(* IEC 61131-3 sources: plc-vscode/tests/st/test-ready/trust-platform/examples/OSCAT/water_booster_pump_station/oop/src, 3 files *)

(* ---- Main.st ---- *)
(* Pattern role: IPump is the contract boundary for the Mediator and Observer example. *)
INTERFACE IPump EXTENDS IComponent
    PROPERTY PumpId : INT
    GET
    END_GET
    END_PROPERTY

    PROPERTY IsHealthy : BOOL
    GET
    END_GET
    END_PROPERTY

    PROPERTY IsRunning : BOOL
    GET
    END_GET
    END_PROPERTY

    PROPERTY RuntimeHours : REAL
    GET
    END_GET
    END_PROPERTY

    PROPERTY SpeedReference : REAL
    GET
    END_GET
    END_PROPERTY

    METHOD Run
    VAR_INPUT
        SpeedReference : REAL;
    END_VAR
    END_METHOD

    METHOD Stop
    END_METHOD
END_INTERFACE

(* Pattern role: IAlarmSubscriber is the contract boundary for the Mediator and Observer example. *)
INTERFACE IAlarmSubscriber
    METHOD OnAlarm
    VAR_INPUT
        ClassId : BYTE;
        Code : DWORD;
        SourceId : INT;
    END_VAR
    END_METHOD
END_INTERFACE

(* Pattern role: PumpDrive is a concrete implementation in the Mediator and Observer example. *)
FUNCTION_BLOCK PumpDrive IMPLEMENTS IPump
VAR
    IdValue : INT;
    FaultValue : BOOL;
    RemoteValue : BOOL := TRUE;
    RunningValue : BOOL;
    RuntimeValue : REAL;
    SpeedValue : REAL;
    ReadyValue : BOOL;
    ErrorValue : BOOL;
    ErrorIdValue : WORD;
    StatusValue : BYTE;
    RuntimeMeter : OntimeMeter;
END_VAR

METHOD PUBLIC Configure
VAR_INPUT
    PumpId : INT;
    RuntimeHoursInitial : REAL;
    Faulted : BOOL;
END_VAR
IdValue := PumpId;
RuntimeValue := RuntimeHoursInitial;
FaultValue := Faulted;
END_METHOD

METHOD PUBLIC Initialize
ReadyValue := TRUE;
RuntimeMeter.Initialize();
RuntimeMeter.Reset();
ClearError();
END_METHOD

METHOD PUBLIC Reset
RunningValue := FALSE;
SpeedValue := REAL#0.0;
ClearError();
END_METHOD

METHOD PUBLIC ClearError
ErrorValue := FALSE;
ErrorIdValue := WORD#0;
StatusValue := BYTE#0;
END_METHOD

METHOD PUBLIC Snapshot : ComponentStatus
VAR
    Result : ComponentStatus;
END_VAR
Result.Ready := ReadyValue;
Result.Error := ErrorValue;
Result.ErrorId := ErrorIdValue;
Result.Status := StatusValue;
Snapshot := Result;
END_METHOD

METHOD PUBLIC Run
VAR_INPUT
    SpeedReference : REAL;
END_VAR
IF NOT FaultValue AND RemoteValue THEN
    RunningValue := TRUE;
    SpeedValue := LIMIT(REAL#0.0, SpeedReference, REAL#100.0);
ELSE
    RunningValue := FALSE;
    SpeedValue := REAL#0.0;
END_IF;
RuntimeMeter.Update(Input := RunningValue);
END_METHOD

METHOD PUBLIC Stop
RunningValue := FALSE;
SpeedValue := REAL#0.0;
RuntimeMeter.Update(Input := FALSE);
END_METHOD

PUBLIC PROPERTY PumpId : INT
GET
    PumpId := IdValue;
END_GET
END_PROPERTY

PUBLIC PROPERTY IsHealthy : BOOL
GET
    IsHealthy := NOT FaultValue AND RemoteValue;
END_GET
END_PROPERTY

PUBLIC PROPERTY IsRunning : BOOL
GET
    IsRunning := RunningValue;
END_GET
END_PROPERTY

PUBLIC PROPERTY RuntimeHours : REAL
GET
    RuntimeHours := RuntimeValue;
END_GET
END_PROPERTY

PUBLIC PROPERTY SpeedReference : REAL
GET
    SpeedReference := SpeedValue;
END_GET
END_PROPERTY

PUBLIC PROPERTY Ready : BOOL
GET
    Ready := ReadyValue;
END_GET
END_PROPERTY

PUBLIC PROPERTY Error : BOOL
GET
    Error := ErrorValue;
END_GET
END_PROPERTY

PUBLIC PROPERTY ErrorId : WORD
GET
    ErrorId := ErrorIdValue;
END_GET
END_PROPERTY

PUBLIC PROPERTY Status : BYTE
GET
    Status := StatusValue;
END_GET
END_PROPERTY
END_FUNCTION_BLOCK

(* Pattern role: HistorianAlarmSubscriber is a concrete implementation in the Mediator and Observer example. *)
FUNCTION_BLOCK HistorianAlarmSubscriber IMPLEMENTS IAlarmSubscriber
VAR
    LastCodeValue : DWORD;
    CountValue : INT;
    Journal : DwordFifo32;
END_VAR

METHOD PUBLIC Initialize
Journal.Initialize();
Journal.Reset();
LastCodeValue := DWORD#0;
CountValue := INT#0;
END_METHOD

METHOD PUBLIC OnAlarm
VAR_INPUT
    ClassId : BYTE;
    Code : DWORD;
    SourceId : INT;
END_VAR
LastCodeValue := Code;
CountValue := CountValue + INT#1;
IF Journal.Push(Value := Code) THEN
END_IF;
END_METHOD

PUBLIC PROPERTY Count : INT
GET
    Count := CountValue;
END_GET
END_PROPERTY

PUBLIC PROPERTY LastCode : DWORD
GET
    LastCode := LastCodeValue;
END_GET
END_PROPERTY
END_FUNCTION_BLOCK

(* Pattern role: MqttAlarmSubscriber is a concrete implementation in the Mediator and Observer example. *)
FUNCTION_BLOCK MqttAlarmSubscriber IMPLEMENTS IAlarmSubscriber
VAR
    PublishReadyValue : BOOL;
    LastCodeValue : DWORD;
END_VAR

METHOD PUBLIC OnAlarm
VAR_INPUT
    ClassId : BYTE;
    Code : DWORD;
    SourceId : INT;
END_VAR
PublishReadyValue := TRUE;
LastCodeValue := Code;
END_METHOD

PUBLIC PROPERTY PublishReady : BOOL
GET
    PublishReady := PublishReadyValue;
END_GET
END_PROPERTY

PUBLIC PROPERTY LastCode : DWORD
GET
    LastCode := LastCodeValue;
END_GET
END_PROPERTY
END_FUNCTION_BLOCK

(* Composition role: AlarmBus owns the collaborating objects used by this Mediator and Observer example. *)
FUNCTION_BLOCK AlarmBus
VAR
    Historian : HistorianAlarmSubscriber;
    Mqtt : MqttAlarmSubscriber;
END_VAR

METHOD PUBLIC Initialize
Historian.Initialize();
END_METHOD

METHOD PUBLIC Publish
VAR_INPUT
    ClassId : BYTE;
    Code : DWORD;
    SourceId : INT;
END_VAR
Historian.OnAlarm(ClassId := ClassId, Code := Code, SourceId := SourceId);
Mqtt.OnAlarm(ClassId := ClassId, Code := Code, SourceId := SourceId);
END_METHOD

PUBLIC PROPERTY HistorianCount : INT
GET
    HistorianCount := Historian.Count;
END_GET
END_PROPERTY

PUBLIC PROPERTY MqttPublishReady : BOOL
GET
    MqttPublishReady := Mqtt.PublishReady;
END_GET
END_PROPERTY
END_FUNCTION_BLOCK

(* Composition role: LeadLagMediator owns the collaborating objects used by this Mediator and Observer example. *)
FUNCTION_BLOCK LeadLagMediator
VAR
    LeadPumpIdValue : INT;
    RunningPumpCountValue : INT;
END_VAR

METHOD PUBLIC Update
VAR_IN_OUT
    Pump1 : PumpDrive;
    Pump2 : PumpDrive;
    Pump3 : PumpDrive;
END_VAR
VAR_INPUT
    DemandLevel : INT;
    SpeedReference : REAL;
END_VAR
VAR
    Lead : IPump;
END_VAR
Pump1.Stop();
Pump2.Stop();
Pump3.Stop();
RunningPumpCountValue := INT#0;

(* Mediator decision: choose the healthy pump with the lowest runtime as lead for wear leveling. *)
IF Pump1.IsHealthy AND (NOT Pump2.IsHealthy OR Pump1.RuntimeHours <= Pump2.RuntimeHours) AND (NOT Pump3.IsHealthy OR Pump1.RuntimeHours <= Pump3.RuntimeHours) THEN
    Lead := Pump1;
ELSIF Pump2.IsHealthy AND (NOT Pump3.IsHealthy OR Pump2.RuntimeHours <= Pump3.RuntimeHours) THEN
    Lead := Pump2;
ELSIF Pump3.IsHealthy THEN
    Lead := Pump3;
ELSE
    LeadPumpIdValue := INT#0;
    RETURN;
END_IF;

LeadPumpIdValue := Lead.PumpId;
Lead.Run(SpeedReference := SpeedReference);
RunningPumpCountValue := INT#1;

IF DemandLevel >= INT#2 THEN
    IF Pump1.IsHealthy AND Pump1.PumpId <> LeadPumpIdValue THEN
        Pump1.Run(SpeedReference := REAL#60.0);
        RunningPumpCountValue := RunningPumpCountValue + INT#1;
    ELSIF Pump2.IsHealthy AND Pump2.PumpId <> LeadPumpIdValue THEN
        Pump2.Run(SpeedReference := REAL#60.0);
        RunningPumpCountValue := RunningPumpCountValue + INT#1;
    ELSIF Pump3.IsHealthy AND Pump3.PumpId <> LeadPumpIdValue THEN
        Pump3.Run(SpeedReference := REAL#60.0);
        RunningPumpCountValue := RunningPumpCountValue + INT#1;
    END_IF;
END_IF;
END_METHOD

PUBLIC PROPERTY LeadPumpId : INT
GET
    LeadPumpId := LeadPumpIdValue;
END_GET
END_PROPERTY

PUBLIC PROPERTY RunningPumpCount : INT
GET
    RunningPumpCount := RunningPumpCountValue;
END_GET
END_PROPERTY
END_FUNCTION_BLOCK

(* Composition role: BoosterStation owns the collaborating objects used by this Mediator and Observer example. *)
FUNCTION_BLOCK BoosterStation
VAR
    Pump1 : PumpDrive;
    Pump2 : PumpDrive;
    Pump3 : PumpDrive;
    Mediator : LeadLagMediator;
    AlarmBusValue : AlarmBus;
    PressureFilter : Pt1Filter;
    Controller : PidController;
    Limits : RealRange;
    Gains : PidGains;
    LeadPumpIdValue : INT;
    RunningPumpCountValue : INT;
    AlarmActiveValue : BOOL;
    CommandValue : REAL;
END_VAR

METHOD PUBLIC Initialize
Pump1.Initialize();
Pump2.Initialize();
Pump3.Initialize();
Pump1.Configure(PumpId := INT#1, RuntimeHoursInitial := REAL#120.0, Faulted := FALSE);
Pump2.Configure(PumpId := INT#2, RuntimeHoursInitial := REAL#20.0, Faulted := FALSE);
Pump3.Configure(PumpId := INT#3, RuntimeHoursInitial := REAL#60.0, Faulted := FALSE);
AlarmBusValue.Initialize();
PressureFilter.Initialize();
PressureFilter.Configure(TimeConstant := T#1s, Gain := REAL#1.0);
Limits.Low := REAL#0.0;
Limits.High := REAL#100.0;
Gains.Kp := REAL#15.0;
Gains.Tn := REAL#1.0;
Gains.Tv := REAL#0.0;
Controller.Initialize();
Controller.Configure(Gains := Gains, Limits := Limits, SupervisionBand := REAL#0.0, Offset := REAL#0.0);
END_METHOD

METHOD PUBLIC SetPumpFaults
VAR_INPUT
    Fault1 : BOOL;
    Fault2 : BOOL;
    Fault3 : BOOL;
END_VAR
Pump1.Configure(PumpId := INT#1, RuntimeHoursInitial := Pump1.RuntimeHours, Faulted := Fault1);
Pump2.Configure(PumpId := INT#2, RuntimeHoursInitial := Pump2.RuntimeHours, Faulted := Fault2);
Pump3.Configure(PumpId := INT#3, RuntimeHoursInitial := Pump3.RuntimeHours, Faulted := Fault3);
END_METHOD

METHOD PUBLIC Update : INT
VAR_INPUT
    StartCommand : BOOL;
    SuctionOk : BOOL;
    HeaderPressure : REAL;
    PressureSetpoint : REAL;
END_VAR
VAR
    FilteredPressure : REAL;
    DemandLevel : INT;
END_VAR
IF NOT SuctionOk THEN
    AlarmActiveValue := TRUE;
    AlarmBusValue.Publish(ClassId := BYTE#1, Code := DWORD#16#A201, SourceId := INT#0);
    Pump1.Stop();
    Pump2.Stop();
    Pump3.Stop();
    (* Suction loss latches lead/running state to zero — pumps are
       commanded stopped, count must reflect that. *)
    RunningPumpCountValue := INT#0;
    LeadPumpIdValue := INT#0;
ELSIF StartCommand THEN
    FilteredPressure := PressureFilter.Update(Sample := HeaderPressure);
    CommandValue := Controller.Update(Actual := FilteredPressure, Target := PressureSetpoint);
    IF PressureSetpoint - FilteredPressure > REAL#1.0 THEN
        DemandLevel := INT#2;
    ELSE
        DemandLevel := INT#1;
    END_IF;
    Mediator.Update(Pump1 := Pump1, Pump2 := Pump2, Pump3 := Pump3, DemandLevel := DemandLevel, SpeedReference := CommandValue);
    LeadPumpIdValue := Mediator.LeadPumpId;
    RunningPumpCountValue := Mediator.RunningPumpCount;
    IF LeadPumpIdValue = INT#0 THEN
        AlarmActiveValue := TRUE;
        AlarmBusValue.Publish(ClassId := BYTE#1, Code := DWORD#16#A202, SourceId := INT#0);
    END_IF;
ELSE
    Pump1.Stop();
    Pump2.Stop();
    Pump3.Stop();
    RunningPumpCountValue := INT#0;
END_IF;
Update := LeadPumpIdValue;
END_METHOD

PUBLIC PROPERTY LeadPumpId : INT
GET
    LeadPumpId := LeadPumpIdValue;
END_GET
END_PROPERTY

PUBLIC PROPERTY RunningPumpCount : INT
GET
    RunningPumpCount := RunningPumpCountValue;
END_GET
END_PROPERTY

PUBLIC PROPERTY AlarmActive : BOOL
GET
    AlarmActive := AlarmActiveValue;
END_GET
END_PROPERTY

PUBLIC PROPERTY HistorianAlarmCount : INT
GET
    HistorianAlarmCount := AlarmBusValue.HistorianCount;
END_GET
END_PROPERTY

PUBLIC PROPERTY MqttPublishReady : BOOL
GET
    MqttPublishReady := AlarmBusValue.MqttPublishReady;
END_GET
END_PROPERTY
END_FUNCTION_BLOCK

(* Scan role: Main wires the example objects and exposes the PLC call path under test. *)
PROGRAM Main
VAR
    Station : BoosterStation;
    StartCommand : BOOL;
    SuctionOk : BOOL;
    Pump1Fault : BOOL;
    Pump2Fault : BOOL;
    Pump3Fault : BOOL;
    HeaderPressureRaw : INT;
    Pump1Enable : BOOL;
    Pump2Enable : BOOL;
    Pump3Enable : BOOL;
    AlarmOut : BOOL;
    HeaderPressure : REAL;
    LeadId : INT;
END_VAR

HeaderPressure := TO_REAL(HeaderPressureRaw) / REAL#100.0;
Station.Initialize();
Station.SetPumpFaults(Fault1 := Pump1Fault, Fault2 := Pump2Fault, Fault3 := Pump3Fault);
LeadId := Station.Update(StartCommand := StartCommand, SuctionOk := SuctionOk, HeaderPressure := HeaderPressure, PressureSetpoint := REAL#4.5);
Pump1Enable := LeadId = INT#1;
Pump2Enable := LeadId = INT#2;
Pump3Enable := LeadId = INT#3;
AlarmOut := Station.AlarmActive;
END_PROGRAM

(* ---- Configuration.st ---- *)
CONFIGURATION WaterBoosterOopConfiguration
RESOURCE Cpu0 ON PLC
    TASK MainTask (INTERVAL := T#100ms, PRIORITY := 1);
    PROGRAM Station WITH MainTask : Main;
END_RESOURCE
VAR_CONFIG
    Station.StartCommand AT %IX0.0 : BOOL;
    Station.SuctionOk AT %IX0.1 : BOOL;
    Station.Pump1Fault AT %IX0.2 : BOOL;
    Station.Pump2Fault AT %IX0.3 : BOOL;
    Station.Pump3Fault AT %IX0.4 : BOOL;
    Station.HeaderPressureRaw AT %IW0 : INT;
    Station.Pump1Enable AT %QX0.0 : BOOL;
    Station.Pump2Enable AT %QX0.1 : BOOL;
    Station.Pump3Enable AT %QX0.2 : BOOL;
    Station.AlarmOut AT %QX0.3 : BOOL;
END_VAR
END_CONFIGURATION

(* ---- Tests.st ---- *)
TEST_PROGRAM BoosterMediatorSelectsLowestRuntimeHealthyPump
VAR
    Station : BoosterStation;
END_VAR

Station.Initialize();
ASSERT_EQUAL(EXPECTED := INT#2, ACTUAL := Station.Update(StartCommand := TRUE, SuctionOk := TRUE, HeaderPressure := REAL#4.0, PressureSetpoint := REAL#4.5));
ASSERT_EQUAL(EXPECTED := INT#2, ACTUAL := Station.LeadPumpId);
ASSERT_EQUAL(EXPECTED := INT#1, ACTUAL := Station.RunningPumpCount);
END_TEST_PROGRAM

TEST_PROGRAM BoosterMediatorFailsOverAndObserverPublishesAlarms
VAR
    Station : BoosterStation;
END_VAR

Station.Initialize();
Station.SetPumpFaults(Fault1 := FALSE, Fault2 := TRUE, Fault3 := FALSE);
ASSERT_EQUAL(EXPECTED := INT#3, ACTUAL := Station.Update(StartCommand := TRUE, SuctionOk := TRUE, HeaderPressure := REAL#4.0, PressureSetpoint := REAL#4.5));

Station.SetPumpFaults(Fault1 := TRUE, Fault2 := TRUE, Fault3 := TRUE);
ASSERT_EQUAL(EXPECTED := INT#0, ACTUAL := Station.Update(StartCommand := TRUE, SuctionOk := TRUE, HeaderPressure := REAL#4.0, PressureSetpoint := REAL#4.5));
ASSERT_TRUE(IN := Station.AlarmActive);
ASSERT_EQUAL(EXPECTED := INT#1, ACTUAL := Station.HistorianAlarmCount);
ASSERT_TRUE(IN := Station.MqttPublishReady);
END_TEST_PROGRAM

(* Multi-cycle observer-fan-out test: drives several alarm-triggering
   scans through one Station and verifies HistorianAlarmCount grows
   monotonically. Catches bugs where the alarm bus re-publishes the
   same event repeatedly, or where the historian counter is reset
   between scans. *)
TEST_PROGRAM BoosterAlarmBusAccumulatesAcrossMultipleEvents
VAR
    Station : BoosterStation;
    InitialHistorian : INT;
END_VAR

Station.Initialize();

(* Scan 1: dry-run condition forces alarm *)
Station.Update(StartCommand := TRUE, SuctionOk := FALSE, HeaderPressure := REAL#4.0, PressureSetpoint := REAL#4.5);
ASSERT_TRUE(IN := Station.AlarmActive);
InitialHistorian := Station.HistorianAlarmCount;
ASSERT_TRUE(IN := InitialHistorian >= INT#1);

(* Scan 2: all pumps faulted forces a different alarm *)
Station.SetPumpFaults(Fault1 := TRUE, Fault2 := TRUE, Fault3 := TRUE);
Station.Update(StartCommand := TRUE, SuctionOk := TRUE, HeaderPressure := REAL#4.0, PressureSetpoint := REAL#4.5);
ASSERT_TRUE(IN := Station.HistorianAlarmCount > InitialHistorian);
ASSERT_TRUE(IN := Station.MqttPublishReady);
END_TEST_PROGRAM

(* Mediator failover regression: pump 2 leads first; when pump 2
   faults, pump 3 takes over within a single same-instance sequence
   (no Initialize between calls). Catches bugs where the mediator
   caches lead selection or fails to re-evaluate fault state. *)
TEST_PROGRAM BoosterMediatorReevaluatesLeadAfterFault
VAR
    Station : BoosterStation;
END_VAR

Station.Initialize();

(* All pumps healthy -> pump 2 leads (lowest runtime) *)
Station.Update(StartCommand := TRUE, SuctionOk := TRUE, HeaderPressure := REAL#4.0, PressureSetpoint := REAL#4.5);
ASSERT_EQUAL(EXPECTED := INT#2, ACTUAL := Station.LeadPumpId);

(* Pump 2 faults -> pump 3 takes lead in the next scan *)
Station.SetPumpFaults(Fault1 := FALSE, Fault2 := TRUE, Fault3 := FALSE);
Station.Update(StartCommand := TRUE, SuctionOk := TRUE, HeaderPressure := REAL#4.0, PressureSetpoint := REAL#4.5);
ASSERT_EQUAL(EXPECTED := INT#3, ACTUAL := Station.LeadPumpId);

(* Pump 2 recovers -> mediator must select a healthy pump (any of 1, 2,
   or 3 is acceptable depending on runtime balance). The point is that
   the mediator re-evaluates rather than caching the previous lead. *)
Station.SetPumpFaults(Fault1 := FALSE, Fault2 := FALSE, Fault3 := FALSE);
Station.Update(StartCommand := TRUE, SuctionOk := TRUE, HeaderPressure := REAL#4.0, PressureSetpoint := REAL#4.5);
ASSERT_TRUE(IN := Station.LeadPumpId >= INT#1);
ASSERT_TRUE(IN := Station.LeadPumpId <= INT#3);
END_TEST_PROGRAM

(* Dry-run permissive: SuctionOk = FALSE blocks all pumps. *)
TEST_PROGRAM BoosterDryRunPermissiveBlocksAllPumps
VAR
    Station : BoosterStation;
END_VAR
Station.Initialize();

(* Suction healthy -> at least one pump runs *)
Station.Update(StartCommand := TRUE, SuctionOk := TRUE, HeaderPressure := REAL#4.0, PressureSetpoint := REAL#4.5);
ASSERT_TRUE(IN := Station.RunningPumpCount >= INT#1);

(* Suction lost -> all pumps must stop, no lead pump *)
Station.Update(StartCommand := TRUE, SuctionOk := FALSE, HeaderPressure := REAL#4.0, PressureSetpoint := REAL#4.5);
ASSERT_EQUAL(EXPECTED := INT#0, ACTUAL := Station.RunningPumpCount);
ASSERT_TRUE(IN := Station.AlarmActive);

(* Suction recovers -> at least one pump runs again (low pressure
   triggers demand). *)
Station.Update(StartCommand := TRUE, SuctionOk := TRUE, HeaderPressure := REAL#4.0, PressureSetpoint := REAL#4.5);
ASSERT_TRUE(IN := Station.RunningPumpCount >= INT#1);
ASSERT_TRUE(IN := Station.LeadPumpId >= INT#1);
END_TEST_PROGRAM

(* StartCommand = FALSE stops all pumps regardless of pressure error. *)
TEST_PROGRAM BoosterStartCommandFalseStopsAllPumps
VAR
    Station : BoosterStation;
END_VAR
Station.Initialize();
Station.Update(StartCommand := TRUE, SuctionOk := TRUE, HeaderPressure := REAL#4.0, PressureSetpoint := REAL#4.5);
ASSERT_TRUE(IN := Station.RunningPumpCount >= INT#1);

(* Stop command -> all pumps stop *)
Station.Update(StartCommand := FALSE, SuctionOk := TRUE, HeaderPressure := REAL#4.0, PressureSetpoint := REAL#4.5);
ASSERT_EQUAL(EXPECTED := INT#0, ACTUAL := Station.RunningPumpCount);
END_TEST_PROGRAM

(* Pressure-on-setpoint case: when pressure == setpoint, no demand. *)
TEST_PROGRAM BoosterAtSetpointHasMinimalDemand
VAR
    Station : BoosterStation;
END_VAR
Station.Initialize();
(* Pressure exactly at setpoint - no error -> minimal pump activity *)
Station.Update(StartCommand := TRUE, SuctionOk := TRUE, HeaderPressure := REAL#4.5, PressureSetpoint := REAL#4.5);
(* Either no pumps or one pump running depending on idle policy *)
ASSERT_TRUE(IN := Station.RunningPumpCount <= INT#1);
END_TEST_PROGRAM

(* Each subscriber observes events independently. *)
TEST_PROGRAM BoosterAlarmBusFansOutToBothSubscribers
VAR
    Station : BoosterStation;
END_VAR
Station.Initialize();

(* Trigger alarm: both Historian count + MQTT flag get set *)
Station.SetPumpFaults(Fault1 := TRUE, Fault2 := TRUE, Fault3 := TRUE);
Station.Update(StartCommand := TRUE, SuctionOk := TRUE, HeaderPressure := REAL#4.0, PressureSetpoint := REAL#4.5);
ASSERT_TRUE(IN := Station.HistorianAlarmCount > INT#0);
ASSERT_TRUE(IN := Station.MqttPublishReady);
END_TEST_PROGRAM

(* Single-pump-fault graceful degradation. *)
TEST_PROGRAM BoosterContinuesWithOnePumpFaulted
VAR
    Station : BoosterStation;
END_VAR
Station.Initialize();
Station.SetPumpFaults(Fault1 := TRUE, Fault2 := FALSE, Fault3 := FALSE);
Station.Update(StartCommand := TRUE, SuctionOk := TRUE, HeaderPressure := REAL#4.0, PressureSetpoint := REAL#4.5);
(* Lead pump is one of the healthy ones (2 or 3) *)
ASSERT_TRUE(IN := (Station.LeadPumpId = INT#2) OR (Station.LeadPumpId = INT#3));
ASSERT_TRUE(IN := Station.LeadPumpId <> INT#1);
END_TEST_PROGRAM

(* Multi-call regression: 20 same-input scans should keep the same lead
   pump selected and not duplicate alarms or recurring publish events
   on healthy operation. *)
TEST_PROGRAM BoosterStableLeadOnHealthyOperation
VAR
    Station : BoosterStation;
    I : INT;
END_VAR
Station.Initialize();
FOR I := 1 TO 20 DO
    Station.Update(StartCommand := TRUE, SuctionOk := TRUE, HeaderPressure := REAL#4.0, PressureSetpoint := REAL#4.5);
END_FOR;
ASSERT_EQUAL(EXPECTED := INT#2, ACTUAL := Station.LeadPumpId);
ASSERT_FALSE(IN := Station.AlarmActive);
ASSERT_EQUAL(EXPECTED := INT#0, ACTUAL := Station.HistorianAlarmCount);
END_TEST_PROGRAM

(* Boundary test: high demand (pressure error >= 1.0) drives the
   mediator to start a lag pump. Total running pumps should be 2. *)
TEST_PROGRAM BoosterHighDemandRunsTwoPumps
VAR
    Station : BoosterStation;
END_VAR
Station.Initialize();
(* Big pressure deficit triggers DemandLevel = 2 (lag pump) *)
Station.Update(StartCommand := TRUE, SuctionOk := TRUE, HeaderPressure := REAL#1.0, PressureSetpoint := REAL#5.0);
ASSERT_EQUAL(EXPECTED := INT#2, ACTUAL := Station.RunningPumpCount);
ASSERT_TRUE(IN := Station.LeadPumpId >= INT#1);
END_TEST_PROGRAM

(* Per-FB isolation: drive a bare PumpDrive object directly and verify
   Run/Stop transitions update IsRunning + SpeedReference. *)
TEST_PROGRAM BoosterPumpDriveStartsAndStopsIndependently
VAR
    Pump : PumpDrive;
END_VAR
Pump.Initialize();
Pump.Configure(PumpId := INT#5, RuntimeHoursInitial := REAL#10.0, Faulted := FALSE);
ASSERT_FALSE(IN := Pump.IsRunning);

Pump.Run(SpeedReference := REAL#75.0);
ASSERT_TRUE(IN := Pump.IsRunning);
ASSERT_NEAR(EXPECTED := REAL#75.0, ACTUAL := Pump.SpeedReference, DELTA := REAL#0.001);

Pump.Stop();
ASSERT_FALSE(IN := Pump.IsRunning);
ASSERT_NEAR(EXPECTED := REAL#0.0, ACTUAL := Pump.SpeedReference, DELTA := REAL#0.001);
END_TEST_PROGRAM

(* Edge input: Run on a faulted pump should not start it; the pump's
   IsHealthy property must gate Run internally. *)
TEST_PROGRAM BoosterPumpDriveRefusesToRunWhenFaulted
VAR
    Pump : PumpDrive;
END_VAR
Pump.Initialize();
Pump.Configure(PumpId := INT#9, RuntimeHoursInitial := REAL#5.0, Faulted := TRUE);
ASSERT_FALSE(IN := Pump.IsHealthy);

Pump.Run(SpeedReference := REAL#80.0);
ASSERT_FALSE(IN := Pump.IsRunning);
ASSERT_NEAR(EXPECTED := REAL#0.0, ACTUAL := Pump.SpeedReference, DELTA := REAL#0.001);
END_TEST_PROGRAM
